FUNCTION_BLOCK "Demo"
{ S7_Optimized_Access := 'TRUE' }
VERSION : 0.1
VAR_INPUT x : DINT; END_VAR
VAR_OUTPUT y : DINT; END_VAR
VAR_IN_OUT a : VARIANT; b : VARIANT; END_VAR
VAR copyDone : BOOL; idx : DINT; END_VAR
BEGIN

#idx := -1; #copyDone := PV_READ(#a, #idx, #b); #y := 0; IF #copyDone THEN #y := 1; END_IF;

END_FUNCTION_BLOCK
